Staubli VAL3: Lab2B_Level2.dtx


